FUNCTION_BLOCK RT_TEST
VAR_INPUT
  CLK : BOOL;
END_VAR
VAR
  r : R_TRIG;
  prevQ : BOOL := FALSE;
END_VAR
BEGIN
  r(CLK := CLK);
  //#ASSERT NOT r.Q : Pbad
END_FUNCTION_BLOCK
